Fanuc KAREL source: NC0016.compact.KL

PROGRAM NC0016
%STACKSIZE=65535
%PRIORITY=65535
%NOLOCKGROUP
ROUTINE R FROM NC0016
ROUTINE R
VAR
S1 : INTEGER
BEGIN
S1=1
IF (S1=1) THEN
S1=(S1 + 2)
ELSE
IF (S1=1) THEN
S1=(S1 + 2)
ELSE
IF (S1=1) THEN
S1=(S1 + 2)
ELSE
IF (S1=1) THEN
S1=(S1 + 2)
ELSE
IF (S1=1) THEN
S1=(S1 + 2)
ELSE
IF (S1=1) THEN
S1=(S1 + 2)
ELSE
IF (S1=1) THEN
S1=(S1 + 2)
ELSE
IF (S1=1) THEN
S1=(S1 + 2)
ELSE
S1=(S1 + 1)
ENDIF
ENDIF
ENDIF
ENDIF
ENDIF
ENDIF
ENDIF
ENDIF
END R
BEGIN
R
END NC0016
